FUNCTION_BLOCK FB_FuseControl_1
VAR_INPUT
	bResetChannels:	BOOL;
END_VAR
VAR_OUTPUT
	fbError:		FB_Error;
END_VAR
VAR
	bInFuse		AT %I* : BOOL;
	bOutFuse	AT %Q* : BOOL;
	
	fbDelay				: TON;
	
	fbRS				: RS;
END_VAR

fbRS(SET := bResetChannels, RESET1 := FALSE);
IF NOT bInFuse THEN
	fbError.M_Set(1, '48V-Sicherung hat ausgelöst', 0, E_ErrorIDs.eFuseTripped, E_ErrorSrcs.eFuse);
	fbDelay(IN := FALSE);
END_IF

IF fbRS.Q1 THEN
	fbDelay(IN := TRUE, PT := T#700MS);
	IF bInFuse THEN
		bOutFuse := TRUE;
	END_IF
	IF fbDelay.Q THEN
		fbDelay(IN := FALSE);
		bOutFuse := FALSE;
		fbRS(SET := bResetChannels, RESET1 := TRUE);
	END_IF
END_IF

END_FUNCTION_BLOCK

(* stored: Version 1.1.0.1, ProductVersion 3.1.4024.12
   POU FB_FuseControl_1: Id {02682e8a-00ae-481b-aba2-dd95afe50c1f}, SpecialFunc None *)
